FUNCTION_BLOCK AOption_OR_2 (* Options-Fan-In: 2 AOption-Sockets IN1/IN2 auf 1 Plug OUT, QI_OUT = IN1 OR IN2. OUT.INIT_CNF geht per E_MUX_2/E_DEMUX_2 an den anfragenden Socket zurueck. Gegenstueck zu AOption_T_2. *)
  (* Standard: 61499-1; Description: Copyright (c) 2026 Meisterschulen am Ostbahnhof This program and the accompanying materials are made available under the terms of the Eclipse Public License 2.0 which is available at https://www.eclipse.org/legal/epl-2.0/ SPDX-License-Identifier: EPL-2.0 *)
  (* Version 1.0, 2026-10-16, Franz Höpfinger, Meisterschulen am Ostbahnhof, E_MUX_2.K merkt den anfragenden Socket, E_DEMUX_2 leitet OUT.INIT_CNF dorthin. Max. 1 offene Anfrage (z.B. hinter einem DEMUX). *)
  PACKAGE Option::merging;
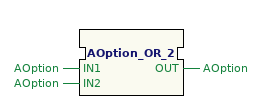
  SOCKETS
    IN1 : Option::AOption; (* Erster AOption-Eingang *)
    IN2 : Option::AOption; (* Zweiter AOption-Eingang *)
  END_SOCKETS
  PLUGS
    OUT : Option::AOption; (* Gemeinsamer Ausgang - aktiv, solange IN1 ODER IN2 aktiv ist *)
  END_PLUGS
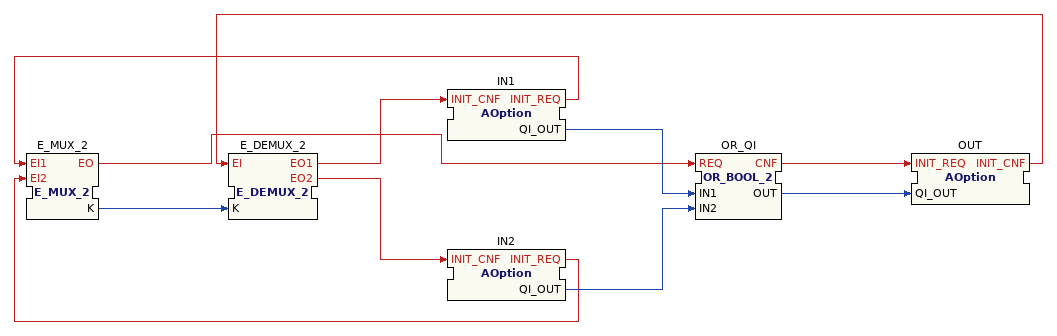
  FBS
    OR_QI : iec61131::booleanOperators::OR_BOOL_2;
    E_MUX_2 : iec61499::events::E_MUX_2;
    E_DEMUX_2 : iec61499::events::E_DEMUX_2;
  END_FBS
  EVENT_CONNECTIONS
    OR_QI.CNF TO OUT.INIT_REQ;
    E_DEMUX_2.EO1 TO IN1.INIT_CNF;
    E_DEMUX_2.EO2 TO IN2.INIT_CNF;
    OUT.INIT_CNF TO E_DEMUX_2.EI;
    IN1.INIT_REQ TO E_MUX_2.EI1;
    IN2.INIT_REQ TO E_MUX_2.EI2;
    E_MUX_2.EO TO OR_QI.REQ;
  END_CONNECTIONS
  DATA_CONNECTIONS
    IN1.QI_OUT TO OR_QI.IN1;
    IN2.QI_OUT TO OR_QI.IN2;
    OR_QI.OUT TO OUT.QI_OUT;
    E_MUX_2.K TO E_DEMUX_2.K;
  END_CONNECTIONS
END_FUNCTION_BLOCK
